(* IEC 61131-3 sources: JingjiangArm/moonboxpro_arm_8.4/Application/Application/任务列表/Main_Task/GNS_MAP/WIDGET, 8 files *)

(* ---- KS_CreatStationIdMap.st ---- *)
(*@CES
Name=KS_CreatStationIdMap
Type=FunctionBlock
TypeGuid=6f9dac99-8de1-4efc-8465-68ac443b7d08
Guid=81839476-edfc-40a3-bf0e-15a9283cc9d6
HasDeclaration=True
HasImplementation=True
*)
{DECLARATION}
FUNCTION KS_CreatStationIdMap : BOOL
(*根据机器类型创建站id的表@根据站号分配表生成*)
(*从1号站开始的|从小到大*)
(*最大128个站*)
VAR_INPUT
	i_iMachineryType	:stEuumMachineryType;(*机器类型@不同设备生成的站列表可能不同*)
	i_piNum				:POINTER TO INT;
	i_paiList			:POINTER TO ARRAY [1..128] OF INT;(*站号从1开始的@总的站列表|需要从小到大*)
	i_piMotionNum		:POINTER TO INT;
	i_paiMotionList		:POINTER TO ARRAY [1..128] OF INT;(*站号从1开始的@运动的站列表|需要从小到大*)
END_VAR
VAR
	(*不同的机型必须要显式赋值*)
	iUnitNum		: INT:=10;(*10色@默认写的是机组式柔印+4压力电机*)
	iLenth			: INT:=128;
	iLenth_Motion	: INT:=128;
	iN				: INT;
	iIndex			: INT;
	iIndex_Motion	: INT;
	iStationId		: INT;
	byStationId		: BYTE;
	aiStationIdList	: ARRAY [1..128] OF INT:=[128(-1)];
	aiMotionStationIdList	: ARRAY [1..128] OF INT:=[128(-1)];
	byTmpL4			: BYTE;
	byTmpH4			: BYTE;
	xStationIdValid	: BOOL;
	xMotionStationIdValid: BOOL;
END_VAR
{IMPLEMENTATION}
iIndex:=0;
iIndex_Motion:=0;
iLenth:=128;
iLenth_Motion:=128;
IF i_paiList<>0 THEN
	iLenth:=SIZEOF(i_paiList^)/SIZEOF(i_paiList^[1]);
END_IF
IF i_paiMotionList<>0 THEN
	iLenth_Motion:=SIZEOF(i_paiMotionList^)/SIZEOF(i_paiMotionList^[1]);
END_IF

CASE i_iMachineryType OF
	MACHINERYTYPE_ROTOGRAVE:;(*凹印*)
	MACHINERYTYPE_FELXO_INLINE,(*机组式柔印*)
	MACHINERYTYPE_FELXO_INLINE_ONEBOTOMROLLER:(*机组式柔印@单底辊*)
		(*不同的机型必须要显式赋值*)
		iUnitNum:=10;
		FOR iN:=1 TO 255 BY 1 DO(*站号最大到255*)
			byStationId:=INT_TO_BYTE(iN);
			byTmpL4:= byStationId AND 16#0F;
			byTmpH4:= SHR(byStationId,4);
			xStationIdValid:=FALSE;
			xMotionStationIdValid:=FALSE;
			IF byTmpL4>0 AND byTmpL4<=iUnitNum THEN(*色组*)
				IF byTmpH4 <= 4 OR(*高4bit小于4是有效的@版辊网辊底辊横向*)
					(byTmpH4 >=7 AND byTmpH4 <= 10)(*压力轴*) THEN
					xStationIdValid:=TRUE;
					IF byTmpH4<>0 THEN(*都是运动的站*)
						xMotionStationIdValid:=TRUE;
					END_IF
				ELSE;
				END_IF
			ELSIF byTmpL4 = 0 THEN(*特殊轴*)
				IF byTmpH4 <= 6 THEN(*高4bit小于6是有效的*)
					xStationIdValid:=TRUE;
					xMotionStationIdValid:=TRUE;
				ELSE;
				END_IF
			ELSE;
			END_IF
			(*再在剩余的里面找找*)
			IF NOT xStationIdValid THEN
				IF byStationId>=92 AND byStationId<=99 THEN
					xStationIdValid:=TRUE;
					xMotionStationIdValid:=TRUE;
				END_IF
			END_IF
			(*所有站*)
			IF xStationIdValid THEN
				iIndex:=iIndex+1;
				IF iIndex<=iLenth THEN
					aiStationIdList[iIndex]:=BYTE_TO_INT(byStationId);
				ELSE
					iIndex:=iLenth;
				END_IF
			END_IF
			(*运动站*)
			IF xMotionStationIdValid THEN
				iIndex_Motion:=iIndex_Motion+1;
				IF iIndex_Motion<=iLenth_Motion THEN
					aiMotionStationIdList[iIndex_Motion]:=BYTE_TO_INT(byStationId);
				ELSE
					iIndex_Motion:=iLenth_Motion;
				END_IF
			END_IF
		END_FOR
	MACHINERYTYPE_FELXO_CL:;(*卫星式柔印*)
	MACHINERYTYPE_OFFSET:;(*胶印机*)
ELSE;
END_CASE

IF i_piNum<>0 THEN
	i_piNum^:=iIndex;
END_IF
IF i_paiList<>0 THEN
	i_paiList^:=aiStationIdList;
END_IF
(*色组站都是不参与运动的|剔除掉*)
IF i_piMotionNum<>0 THEN
	i_piMotionNum^:=iIndex_Motion;
END_IF
IF i_paiMotionList<>0 THEN
	i_paiMotionList^:=aiMotionStationIdList;
END_IF

KS_CreatStationIdMap:=iIndex<>0;

(* ---- KS_GetAxisInfByStationIdForMap.st ---- *)
(*@CES
Name=KS_GetAxisInfByStationIdForMap
Type=FunctionBlock
TypeGuid=6f9dac99-8de1-4efc-8465-68ac443b7d08
Guid=05eda7a9-c666-455e-82aa-6ccc3756d356
HasDeclaration=True
HasImplementation=True
*)
{DECLARATION}
FUNCTION KS_GetAxisInfByStationIdForMap : stEnumAxisId
(*通过站号id获取轴信息@依赖定义的站号配置表(一般不会变化)*)
(*不处理0号站*)
VAR_INPUT
	i_iStationId:INT;(*站号*)
	i_piFuncId:POINTER TO stEnumFuncId;(*只针对色组轴*)
	i_piMoveType:POINTER TO stEnumMoveType;(*运动的类型也可以获取*)
END_VAR
VAR
	iAxisId		: stEnumAxisId		:=AXISID_INVALID;
	iFuncId		: stEnumFuncId		:=FUNCID_NULL;(*只针对色组轴*)
	iMoveType	: stEnumMoveType	:=MOVETYPE_NULL;(*运动的类型也可以获取*)
	byStationId	: BYTE;
	byTmpL4		: BYTE;(*低4bit*)
	byTmpH4		: BYTE;(*高4bit*)
	//ilen:int;
END_VAR
{IMPLEMENTATION}
IF i_iStationId>0 AND i_iStationId<=255 THEN
	byStationId:=INT_TO_BYTE(i_iStationId);
	byTmpL4:= byStationId AND 16#0F;
	byTmpH4:= SHR(byStationId,4);
	(*检查是不是色组@按照规则低4位为色组id号*)
	IF byTmpL4>0 AND byTmpL4<=16#0F THEN
		//iAxisId := iTmpL4;(*和枚举定义对应*)
		//ilen := SIZEOF(iAxisId);
		KS_Int2Enum(ADR(iAxisId),BYTE_TO_INT(byTmpL4)(*iTmpL4*));
		(*高bit代表功能*)
		CASE byTmpH4 OF
			0:iFuncId:=FUNCID_CONTROL;					iMoveType:=MOVETYPE_NULL;
			1:iFuncId:=FUNCID_PRNROLLER;				iMoveType:=MOVETYPE_ROTARY_SUPERPOS;
			2:iFuncId:=FUNCID_NETROLLER;				iMoveType:=MOVETYPE_ROTARY;
			3:iFuncId:=FUNCID_BOTTOMROLLER;				iMoveType:=MOVETYPE_ROTARY;
			4:iFuncId:=FUNCID_HORZ;						iMoveType:=MOVETYPE_TRAP;
			5:(*不是色组轴*)iAxisId:=AXISID_INVALID;
			6:(*不是色组轴*)iAxisId:=AXISID_INVALID;
			7:iFuncId:=FUNCID_PRNROLLER_PRESSURE_M;		iMoveType:=MOVETYPE_GANTRY;
			8:iFuncId:=FUNCID_PRNROLLER_PRESSURE_G;		iMoveType:=MOVETYPE_GANTRY;
			9:iFuncId:=FUNCID_NETROLLER_PRESSURE_M;		iMoveType:=MOVETYPE_GANTRY;
			10:iFuncId:=FUNCID_NETROLLER_PRESSURE_G;	iMoveType:=MOVETYPE_GANTRY;
		ELSE;
		END_CASE
	ELSIF byTmpL4=0 THEN(*低位为0|主要收放牵和收放料*)
		CASE byTmpH4 OF
			1:(*放A*)	iAxisId:=AXISID_UWA;				iMoveType:=MOVETYPE_ROTARY;
			2:(*放B*)	iAxisId:=AXISID_UWB;				iMoveType:=MOVETYPE_ROTARY;
			3:(*收A*)	iAxisId:=AXISID_RWA;				iMoveType:=MOVETYPE_ROTARY;
			4:(*收B*)	iAxisId:=AXISID_RWB;				iMoveType:=MOVETYPE_ROTARY;
			5:(*放牵*)	iAxisId:=AXISID_IF;					iMoveType:=MOVETYPE_ROTARY;
			6:(*收牵*)	iAxisId:=AXISID_OF;					iMoveType:=MOVETYPE_ROTARY;
		ELSE;
		END_CASE
	ELSE;
	END_IF

	(*还有剩余的双收双放应用到的站处理|这部分就单独处理吧*)
	IF iAxisId = AXISID_INVALID THEN(*未找到就再找找*)
		CASE byStationId OF
			92:(*放A@II*)iAxisId:=AXISID_UWA_II;				iMoveType:=MOVETYPE_ROTARY;
			93:(*放B@II*)iAxisId:=AXISID_UWB_II;				iMoveType:=MOVETYPE_ROTARY;
			94:(*收A@II*)iAxisId:=AXISID_RWA_II;				iMoveType:=MOVETYPE_ROTARY;
			95:(*收B@II*)iAxisId:=AXISID_RWB_II;				iMoveType:=MOVETYPE_ROTARY;
			96:(*收牵*);
			97:(*放牵@II*)iAxisId:=AXISID_IF_II;				iMoveType:=MOVETYPE_ROTARY;
			98:(*收牵@II*)iAxisId:=AXISID_OF_II;				iMoveType:=MOVETYPE_ROTARY;
			99:(*中心辊*)iAxisId:=AXISID_CENTER;				iMoveType:=MOVETYPE_ROTARY;
		ELSE;
		END_CASE
	END_IF
END_IF
IF i_piFuncId<>0 THEN
	i_piFuncId^:=iFuncId;
END_IF
IF i_piMoveType<>0 THEN
	i_piMoveType^:=iMoveType;
END_IF

KS_GetAxisInfByStationIdForMap:=iAxisId;

(* ---- KS_GetLogicAxisInfByStationIdForMap.st ---- *)
(*@CES
Name=KS_GetLogicAxisInfByStationIdForMap
Type=FunctionBlock
TypeGuid=6f9dac99-8de1-4efc-8465-68ac443b7d08
Guid=2d4d40f4-a928-4a47-8c3c-7c3d2312de1c
HasDeclaration=True
HasImplementation=True
*)
{DECLARATION}
FUNCTION KS_GetLogicAxisInfByStationIdForMap : INT(*返回逻辑轴id*)
(*通过站号获取逻辑轴信息@轴号和核号|基于xml文件*)
(*实际站号后面都是叠加轴*)
VAR_INPUT
	i_iStationId			:INT;
	i_iMachineryType		:stEuumMachineryType;(*机器类型@不同设备生成的站列表可能不同*)
	(*根据xml配置表获得*)
	i_piCoreId				:POINTER TO INT;(*核id*)
	i_piLogicAxisIdSuperPos	:POINTER TO INT;(*叠加轴id*)
END_VAR
VAR
	iN:INT;
	iStationIdTmp: INT;(*站id*)
	iCoreId: INT:=-1;(*核id*)
	iLogicAxisId:INT:=-1;(*逻辑轴id*)
	iLogicAxisIdSuperPos:INT:=-1;(*叠加轴id*)
	(*不同的机型必须要显式赋值*)
	(*色组数@默认写的是机组式柔印+4压力电机*)
	iUnitNum:INT:=10;
	(*核1核2分配的站个数@默认写的是机组式柔印+4压力电机*)
	byStationNum_Core1: BYTE:=53;
	byStationNum_Core2: BYTE:=40;
	iMoveStationNum: INT:=0;(*运动站个数*)
	aiMoveStationIdList: ARRAY [1..128] OF INT;(*运动站id列表*)
	aiStationIdListTmp: ARRAY [1..128] OF INT;
	iMachineryType: stEuumMachineryType;
	iLogicAxisSaIdCalcSuperAxisId: INT;(*计算叠加轴id时逻辑轴起始@不包含*)
	iLogicAxisEdIdCalcSuperAxisId: INT;(*计算叠加轴id时逻辑轴结束@包含*)
END_VAR
{IMPLEMENTATION}
IF i_iStationId>0 AND i_iStationId<=255 THEN
	iMachineryType:=i_iMachineryType;
	(*生成合理的运动站号表@该表和core1 2的逻辑轴id是有对应关系的@xml文件*)
	KS_CreatStationIdMap(iMachineryType,0, 0, ADR(iMoveStationNum), ADR(aiMoveStationIdList));
	CASE iMachineryType OF
		MACHINERYTYPE_ROTOGRAVE:;(*凹印*)
		MACHINERYTYPE_FELXO_INLINE,(*机组式柔印*)
		MACHINERYTYPE_FELXO_INLINE_ONEBOTOMROLLER:(*机组式柔印@单底辊*)
			(*不同的机型必须要显式赋值*)
			iUnitNum:=10;(*4电机压力限制最大只能10色*)
			byStationNum_Core1:=53;(*核1的实际站个数*)
			byStationNum_Core2:=40;(*核2的实际站个数*)
			(*把核1的站id取出来*)
			SysMemCpy(ADR(aiStationIdListTmp),
					ADR(aiMoveStationIdList),
					SIZEOF(aiMoveStationIdList[1])*byStationNum_Core1);
			FOR iN:=1 TO byStationNum_Core1 BY 1 DO
				iStationIdTmp:=aiStationIdListTmp[iN];
				IF iStationIdTmp = i_iStationId THEN
					iCoreId:=1;
					iLogicAxisId:=iN;
					(*叠加轴处理*)
					IF iMachineryType = MACHINERYTYPE_FELXO_INLINE_ONEBOTOMROLLER THEN
						(*默认的套色轴是底辊*)
						iLogicAxisSaIdCalcSuperAxisId:=(iUnitNum+1)*2+1;
						iLogicAxisEdIdCalcSuperAxisId:=(iUnitNum+1)*3;
					ELSE(*默认套色轴是在版辊*)
						iLogicAxisSaIdCalcSuperAxisId:=1;
						iLogicAxisEdIdCalcSuperAxisId:=iUnitNum+1;
					END_IF

					IF iN>iLogicAxisSaIdCalcSuperAxisId AND
						iN<=iLogicAxisEdIdCalcSuperAxisId THEN
						(*eg:1色版辊叠加轴;iN:=2, 叠加id=53 + 2 - 1 = 54*)
						(*eg:1色底辊叠加轴;iN:=24, 叠加id=53 + 24 - 23 = 54*)
						iLogicAxisIdSuperPos:=BYTE_TO_INT(byStationNum_Core1) + iN - iLogicAxisSaIdCalcSuperAxisId;
					END_IF
					EXIT;
				END_IF
			END_FOR

			IF iCoreId = -1 THEN(*未找到,继续找*)
				(*把核2的站id取出来*)
				SysMemSet(ADR(aiStationIdListTmp),0,SIZEOF(aiStationIdListTmp));
				SysMemCpy(ADR(aiStationIdListTmp),
						ADR(aiMoveStationIdList[byStationNum_Core1+1]),
						SIZEOF(aiMoveStationIdList[1])*byStationNum_Core2);

				FOR iN:=1 TO byStationNum_Core2 BY 1 DO
					iStationIdTmp:=aiStationIdListTmp[iN];
					IF iStationIdTmp = i_iStationId THEN
						iCoreId:=2;
						iLogicAxisId:=iN;
						(*叠加轴处理*)
						IF iN<=iUnitNum THEN
							(*eg:1色版辊M侧压力电机龙门叠加轴;iN:=1, 叠加id= 40 + 1 = 41*)
							iLogicAxisIdSuperPos:=BYTE_TO_INT(byStationNum_Core2) + iN;
						ELSIF iN>iUnitNum*3 THEN(*网辊M侧@不需要处理叠加轴*);
						ELSIF iN>iUnitNum*2 THEN(*再偏移一个版辊G侧压力电机|是网辊M侧的索引*)
							(*eg:1色网辊M侧压力电机龙门叠加轴;iN:=21, 叠加id= 40 + 21 - 10 = 51*)
							iLogicAxisIdSuperPos:=BYTE_TO_INT(byStationNum_Core2) + iN - iUnitNum;
						END_IF
						EXIT;
					END_IF
				END_FOR
			END_IF
		MACHINERYTYPE_FELXO_CL:;(*卫星式柔印*)
		MACHINERYTYPE_OFFSET:;(*胶印机*)
	ELSE;
	END_CASE
ELSE;
END_IF

IF i_piCoreId<>0 THEN
	i_piCoreId^:=iCoreId;
END_IF
IF i_piLogicAxisIdSuperPos<>0 THEN
	i_piLogicAxisIdSuperPos^:=iLogicAxisIdSuperPos;
END_IF
KS_GetLogicAxisInfByStationIdForMap:=iLogicAxisId;

(* ---- KS_GetStationInf.st ---- *)
(*@CES
Name=KS_GetStationInf
Type=FunctionBlock
TypeGuid=6f9dac99-8de1-4efc-8465-68ac443b7d08
Guid=b7f0280a-edd9-42bd-a20b-0c2dea9f3ec3
HasDeclaration=True
HasImplementation=True
*)
{DECLARATION}
FUNCTION KS_GetStationInf : BOOL
(*获取站的信息*)
VAR_INPUT
	i_iStationId			: INT;
	i_pstStationInf			: POINTER TO StStationInf;
	i_pstStSysStationInf	: POINTER TO StSysStationInf;
END_VAR
VAR
	iN: INT;
	pstStationInf				: POINTER TO StStationInf;
	xFindIt: BOOL;
END_VAR

{IMPLEMENTATION}
KS_InitStationInf(i_pstStationInf);
IF i_iStationId>0 AND i_iStationId<=255 THEN
	FOR iN:=1 TO i_pstStSysStationInf^.byStationNum BY 1 DO
		pstStationInf:=ADR(i_pstStSysStationInf^.astStationInf[iN]);
		IF pstStationInf^.xValid THEN(*信息有效了*)
			IF pstStationInf^.iStationId = i_iStationId THEN
				xFindIt:=TRUE;
				EXIT;
			END_IF
		END_IF
	END_FOR

	(*结构体初始化*)
	IF xFindIt THEN
		i_pstStationInf^:=pstStationInf^;
	END_IF
END_IF
KS_GetStationInf:=xFindIt;

(* ---- KS_InitGantryAxisInf.st ---- *)
(*@CES
Name=KS_InitGantryAxisInf
Type=FunctionBlock
TypeGuid=6f9dac99-8de1-4efc-8465-68ac443b7d08
Guid=ab05e6d0-ef39-4b76-beb4-016762606a5a
HasDeclaration=True
HasImplementation=True
*)
{DECLARATION}
FUNCTION KS_InitGantryAxisInf : BOOL
VAR_INPUT
	i_pstStGantryAxisInf :POINTER TO StGantryAxisInf;
END_VAR
VAR
	stStGantryAxisInf :StGantryAxisInf:=(
								iAxisId:=-1,(*色组号*)
								iFuncId:=FUNCID_NULL,(*版辊\网纹辊*)
								iCoreId:=-1,(*核id*)
								iLogicAxisId_M:=-1,(*操作侧逻辑轴id*)
								iLogicAxisId_G:=-1,(*操作侧逻辑轴id*)
								iLogicAxisId_SuperPos:=-1);
END_VAR
{IMPLEMENTATION}
IF i_pstStGantryAxisInf<>0 THEN
	i_pstStGantryAxisInf^:=stStGantryAxisInf;
END_IF

(* ---- KS_InitStationInf.st ---- *)
(*@CES
Name=KS_InitStationInf
Type=FunctionBlock
TypeGuid=6f9dac99-8de1-4efc-8465-68ac443b7d08
Guid=78672f31-3286-4bff-bedb-6c7e7d7440a9
HasDeclaration=True
HasImplementation=True
*)
{DECLARATION}
FUNCTION KS_InitStationInf : BOOL
(*初始化结构体*)
VAR_INPUT
	i_pstInf:POINTER TO StStationInf;
END_VAR
VAR
	stInf:StStationInf:=(xValid:=FALSE,
						iAxisId:=AXISID_INVALID,
						iStationId:=-1,
						iFuncId:=FUNCID_NULL,
						iMoveType:=MOVETYPE_NULL,
						udiStationType:=0,
						iCoreId_LogicAxis:=-1,
						iCoreId_LogicAxisSuperPos:=-1,
						iLogicAxisId:=-1,
						iLogicAxisIdSuperPos:=-1,
						xRemoteEncValid:=FALSE,
						iRemoteSrcId:=-1);
END_VAR
{IMPLEMENTATION}
IF i_pstInf<>0 THEN
	i_pstInf^:=stInf;
END_IF

(* ---- KS_Int2Enum.st ---- *)
(*@CES
Name=KS_Int2Enum
Type=FunctionBlock
TypeGuid=6f9dac99-8de1-4efc-8465-68ac443b7d08
Guid=ce208212-85df-4d43-9cce-e1a5fdafda9b
HasDeclaration=True
HasImplementation=True
*)
{DECLARATION}
FUNCTION KS_Int2Enum : BOOL
//枚举类型按照2个字节处理@简单点
VAR_INPUT
	i_stEnumAdr:DWORD;//枚举地址
	i_iData:INT;//转换值
END_VAR
VAR
	pitmp:POINTER TO INT;
END_VAR

{IMPLEMENTATION}
IF i_stEnumAdr<>0 THEN
	pitmp := i_stEnumAdr;
	pitmp^:= i_iData;
END_IF

(* ---- KS_IsUnitAxisId.st ---- *)
(*@CES
Name=KS_IsUnitAxisId
Type=FunctionBlock
TypeGuid=6f9dac99-8de1-4efc-8465-68ac443b7d08
Guid=fbe75c62-94e0-460b-970c-a4df6e13b71e
HasDeclaration=True
HasImplementation=True
*)
{DECLARATION}
FUNCTION KS_IsUnitAxisId : BOOL
(*色组轴id@轴id枚举里包含了非色组轴的定义*)
VAR_INPUT
	i_iAxisId:stEnumAxisId;
END_VAR
VAR
	xResult: BOOL;
END_VAR
{IMPLEMENTATION}
IF i_iAxisId>=AXISID_1U AND
	i_iAxisId<=AXISID_15U THEN
	xResult:=TRUE;
END_IF
KS_IsUnitAxisId:=xResult;
